Fanuc KAREL source: KT00431.KL

PROGRAM KT00431
%NOLOCKGROUP
VAR
  P1: JOINTPOS
  P2: POSITION
  OUT: BOOLEAN
BEGIN
  OUT = P1 > P2
END KT00431
